(* PLC project g_ton_single, Anonymous Benchmark Suite 1.0 *)
(* stored: creationDateTime 2026-08-26T00:00:00 *)

PROGRAM g_ton_single
  VAR_INPUT
    Btn : BOOL;
  END_VAR
  VAR_OUTPUT
    Light : BOOL;
  END_VAR
  VAR
    TON0 : TON;
  END_VAR

(* LD diagram, written out as Structured Text *)
TON0(IN := Btn, PT := T#30ms);
Light := TON0.Q;
END_PROGRAM

CONFIGURATION Config0
  RESOURCE Res0 ON PLC
    TASK tcyclic(INTERVAL := T#10ms, PRIORITY := 0);
    PROGRAM inst0 WITH tcyclic : g_ton_single;
  END_RESOURCE
END_CONFIGURATION
